// Mitsubishi GX Works2 project: 수위제어2   PLC: Q02/Q02H

PROGRAM MAIN
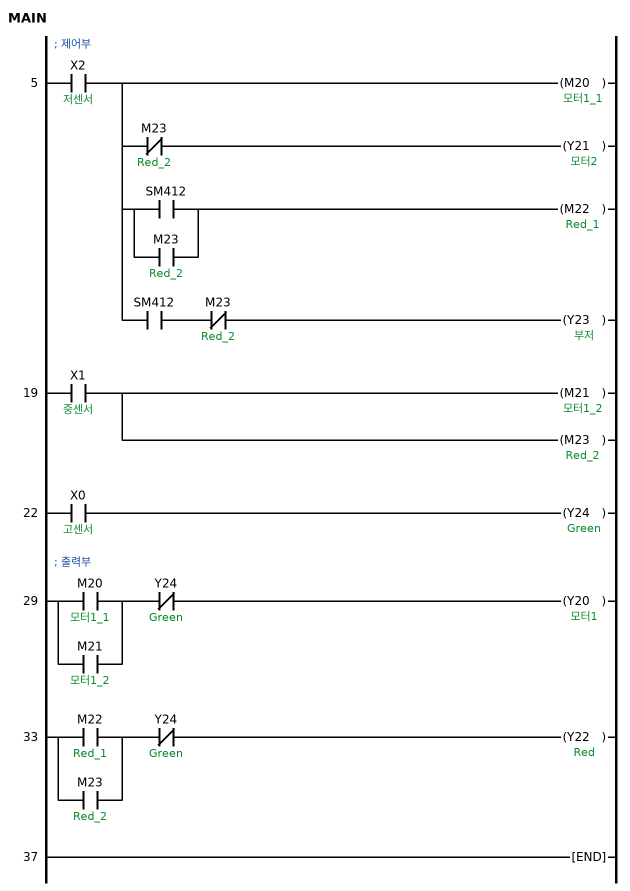
; 제어부
5     LD      X2  ; 저센서
      OUT     M20  ; 모터1_1
      MPS
      ANI     M23  ; Red_2
      OUT     Y21  ; 모터2
      MRD
      LD      SM412
      OR      M23  ; Red_2
      ANB
      OUT     M22  ; Red_1
      MPP
      AND     SM412
      ANI     M23  ; Red_2
      OUT     Y23  ; 부저
19    LD      X1  ; 중센서
      OUT     M21  ; 모터1_2
      OUT     M23  ; Red_2
22    LD      X0  ; 고센서
      OUT     Y24  ; Green
; 출력부
29    LD      M20  ; 모터1_1
      OR      M21  ; 모터1_2
      ANI     Y24  ; Green
      OUT     Y20  ; 모터1
33    LD      M22  ; Red_1
      OR      M23  ; Red_2
      ANI     Y24  ; Green
      OUT     Y22  ; Red
37    END
END_PROGRAM

// device comments not shown above
X3  ; 테스트
